(* IEC 61131-3 sources: PLCHaT-dataset/benchmark_mutated/253_AlarmProcess/mutation_1/syntax_check, 1 file *)

(* ---- 253_AlarmProcess.st.clean.st ---- *)
FUNCTION_BLOCK AlarmProcess
VAR_INPUT
    Value : REAL;
    hiLevel : REAL;
    loLevel : REAL;
    hystWindow : REAL;
END_VAR
VAR_OUTPUT
    hiAlarm : BOOL;
    loAlarm : BOOL;
    error : BOOL;
    status : WORD;
END_VAR
VAR
    tempStatus : WORD;
END_VAR

error := FALSE;
tempStatus := 0;

IF loLevel >= hiLevel THEN
    error := TRUE;
    tempStatus := 16#8001;
ELSIF hystWindow >= (hiLevel - loLevel) THEN
    error := FALSE;
    tempStatus := 16#0000;
ELSE
    IF Value > hiLevel THEN
        hiAlarm := TRUE;
    ELSIF Value < (hiLevel - hystWindow) THEN
        hiAlarm := FALSE;
    END_IF;

    IF Value < loLevel THEN
        loAlarm := TRUE;
    ELSIF Value > (loLevel + hystWindow) THEN
        loAlarm := FALSE;
    END_IF;
END_IF;

status := tempStatus;

END_FUNCTION_BLOCK
